TYPE ST_PolarIIChamber_CupServiceStatus :
STRUCT
	Lift : ST_PolarIIChamber_CupLiftServiceStatus;
	Drainer : ST_PolarIIChamber_SelectThreeServiceStatus;
END_STRUCT
END_TYPE

(* stored: Version 1.1.0.1, ProductVersion 3.1.4026.18
   DUT ST_PolarIIChamber_CupServiceStatus: Id {14000000-0000-0000-0000-000000000063} *)
